FUNCTION_BLOCK DesidratacaoLodo_HMI (* Service Interface Function Block Type *)
  (* Standard: 61499-2 *)
  (* Version 1.2, 21/10/2026, Hidryco, Hidryco, IHM da DesidratacaoLodo 1.2: rodizio e PID nos sub-CATs Revezamento e PID *)
  PACKAGE Hidryco.HidrycoLib;
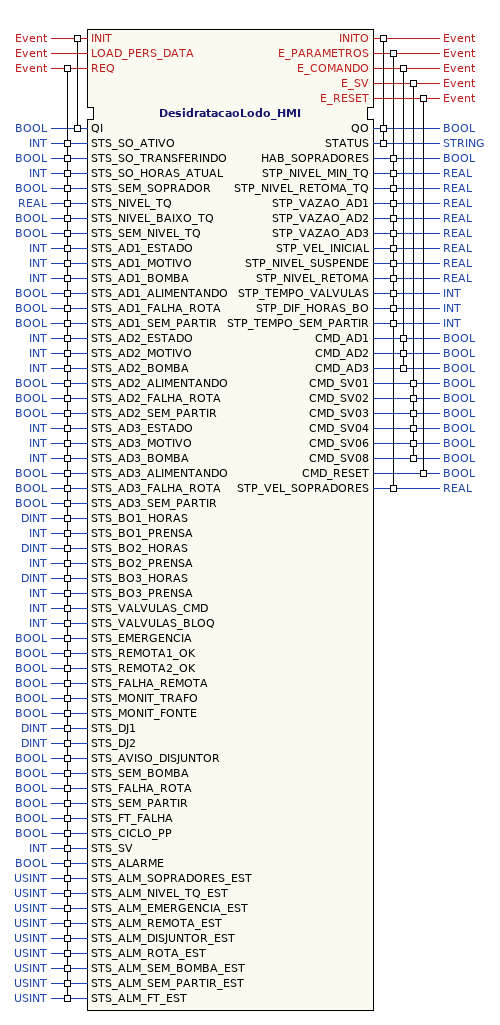
  EVENT_INPUT
    INIT WITH QI;
    LOAD_PERS_DATA; (* Reenvia os parametros persistentes *)
    REQ WITH STS_SO_ATIVO, STS_SO_TRANSFERINDO, STS_SO_HORAS_ATUAL, STS_SEM_SOPRADOR, STS_NIVEL_TQ, STS_NIVEL_BAIXO_TQ, STS_SEM_NIVEL_TQ, STS_AD1_ESTADO, STS_AD1_MOTIVO, STS_AD1_BOMBA, STS_AD1_ALIMENTANDO, STS_AD1_FALHA_ROTA, STS_AD1_SEM_PARTIR, STS_AD2_ESTADO, STS_AD2_MOTIVO, STS_AD2_BOMBA, STS_AD2_ALIMENTANDO, STS_AD2_FALHA_ROTA, STS_AD2_SEM_PARTIR, STS_AD3_ESTADO, STS_AD3_MOTIVO, STS_AD3_BOMBA, STS_AD3_ALIMENTANDO, STS_AD3_FALHA_ROTA, STS_AD3_SEM_PARTIR, STS_BO1_HORAS, STS_BO1_PRENSA, STS_BO2_HORAS, STS_BO2_PRENSA, STS_BO3_HORAS, STS_BO3_PRENSA, STS_VALVULAS_CMD, STS_VALVULAS_BLOQ, STS_EMERGENCIA, STS_REMOTA1_OK, STS_REMOTA2_OK, STS_FALHA_REMOTA, STS_MONIT_TRAFO, STS_MONIT_FONTE, STS_DJ1, STS_DJ2, STS_AVISO_DISJUNTOR, STS_SEM_BOMBA, STS_FALHA_ROTA, STS_SEM_PARTIR, STS_FT_FALHA, STS_CICLO_PP, STS_SV, STS_ALARME, STS_ALM_SOPRADORES_EST, STS_ALM_NIVEL_TQ_EST, STS_ALM_EMERGENCIA_EST, STS_ALM_REMOTA_EST, STS_ALM_DISJUNTOR_EST, STS_ALM_ROTA_EST, STS_ALM_SEM_BOMBA_EST, STS_ALM_SEM_PARTIR_EST, STS_ALM_FT_EST; (* Atualizacao de status *)
  END_EVENT
  EVENT_OUTPUT
    INITO WITH QO, STATUS;
    E_PARAMETROS WITH HAB_SOPRADORES, STP_NIVEL_MIN_TQ, STP_NIVEL_RETOMA_TQ, STP_VAZAO_AD1, STP_VAZAO_AD2, STP_VAZAO_AD3, STP_VEL_INICIAL, STP_NIVEL_SUSPENDE, STP_NIVEL_RETOMA, STP_TEMPO_VALVULAS, STP_DIF_HORAS_BO, STP_TEMPO_SEM_PARTIR, STP_VEL_SOPRADORES;
    E_COMANDO WITH CMD_AD1, CMD_AD2, CMD_AD3;
    E_SV WITH CMD_SV01, CMD_SV02, CMD_SV03, CMD_SV04, CMD_SV06, CMD_SV08;
    E_RESET WITH CMD_RESET;
  END_EVENT
  VAR_INPUT
    QI : BOOL;
    STS_SO_ATIVO : INT; (* Soprador designado: 0 nenhum, 1 SO-01, 2 SO-02 *)
    STS_SO_TRANSFERINDO : BOOL; (* Rodizio em andamento (os dois ligados) *)
    STS_SO_HORAS_ATUAL : INT; (* Horas do soprador atual desde a ultima troca *)
    STS_SEM_SOPRADOR : BOOL; (* Automatico sem nenhum soprador disponivel (risco de sedimentacao) *)
    STS_NIVEL_TQ : REAL; (* Nivel usado no intertravamento (maior entre LIT-01 e LIT-02 validos, %) *)
    STS_NIVEL_BAIXO_TQ : BOOL; (* Tanques de estocagem em nivel baixo: bombas suspensas *)
    STS_SEM_NIVEL_TQ : BOOL; (* LIT-01 e LIT-02 em falha: bombas suspensas *)
    STS_AD1_ESTADO : INT; (* AD-01: 0 parado, 1 abrindo valvulas, 2 partindo bomba, 3 alimentando, 4 suspenso, 5 parando *)
    STS_AD1_MOTIVO : INT; (* AD-01: 0 ok, 1 prensa indisponivel, 2 setpoint zero, 3 sem bomba ou rota, 4 houve falha de rota, 5 emergencia, 6 floculador cheio, 7 tanque baixo, 8 FT em falha, 9 prensa nao partiu *)
    STS_AD1_BOMBA : INT; (* AD-01: bomba em uso (0 nenhuma, 1 a 3 = BO-01 a BO-03) *)
    STS_AD1_ALIMENTANDO : BOOL; (* AD-01 sendo alimentada *)
    STS_AD1_FALHA_ROTA : BOOL; (* AD-01: valvula da rota nao abriu/fechou ou saiu de posicao com a bomba em uso (memorizado; outra rota e tentada) *)
    STS_AD1_SEM_PARTIR : BOOL; (* AD-01 alimentada e a prensa nao partiu no tempo *)
    STS_AD2_ESTADO : INT; (* AD-02: 0 parado, 1 abrindo valvulas, 2 partindo bomba, 3 alimentando, 4 suspenso, 5 parando *)
    STS_AD2_MOTIVO : INT; (* AD-02: 0 ok, 1 prensa indisponivel, 2 setpoint zero, 3 sem bomba ou rota, 4 houve falha de rota, 5 emergencia, 6 floculador cheio, 7 tanque baixo, 8 FT em falha, 9 prensa nao partiu *)
    STS_AD2_BOMBA : INT; (* AD-02: bomba em uso (0 nenhuma, 1 a 3 = BO-01 a BO-03) *)
    STS_AD2_ALIMENTANDO : BOOL; (* AD-02 sendo alimentada *)
    STS_AD2_FALHA_ROTA : BOOL; (* AD-02: valvula da rota nao abriu/fechou ou saiu de posicao com a bomba em uso (memorizado; outra rota e tentada) *)
    STS_AD2_SEM_PARTIR : BOOL; (* AD-02 alimentada e a prensa nao partiu no tempo *)
    STS_AD3_ESTADO : INT; (* AD-03: 0 parado, 1 abrindo valvulas, 2 partindo bomba, 3 alimentando, 4 suspenso, 5 parando *)
    STS_AD3_MOTIVO : INT; (* AD-03: 0 ok, 1 prensa indisponivel, 2 setpoint zero, 3 sem bomba ou rota, 4 houve falha de rota, 5 emergencia, 6 floculador cheio, 7 tanque baixo, 8 FT em falha, 9 prensa nao partiu *)
    STS_AD3_BOMBA : INT; (* AD-03: bomba em uso (0 nenhuma, 1 a 3 = BO-01 a BO-03) *)
    STS_AD3_ALIMENTANDO : BOOL; (* AD-03 sendo alimentada *)
    STS_AD3_FALHA_ROTA : BOOL; (* AD-03: valvula da rota nao abriu/fechou ou saiu de posicao com a bomba em uso (memorizado; outra rota e tentada) *)
    STS_AD3_SEM_PARTIR : BOOL; (* AD-03 alimentada e a prensa nao partiu no tempo *)
    STS_BO1_HORAS : DINT; (* BO-01: horas de operacao (rodizio) *)
    STS_BO1_PRENSA : INT; (* BO-01: prensa atendida (0 nenhuma, 1 a 3) *)
    STS_BO2_HORAS : DINT; (* BO-02: horas de operacao (rodizio) *)
    STS_BO2_PRENSA : INT; (* BO-02: prensa atendida (0 nenhuma, 1 a 3) *)
    STS_BO3_HORAS : DINT; (* BO-03: horas de operacao (rodizio) *)
    STS_BO3_PRENSA : INT; (* BO-03: prensa atendida (0 nenhuma, 1 a 3) *)
    STS_VALVULAS_CMD : INT; (* Valvulas do barrilete comandadas abertas (bit 0 = VA-06 ... bit 7 = VA-13) *)
    STS_VALVULAS_BLOQ : INT; (* Valvulas do barrilete bloqueadas por falha de rota ate o reset (bit 0 = VA-06 ... bit 7 = VA-13) *)
    STS_EMERGENCIA : BOOL; (* Emergencia do PCM LODO acionada *)
    STS_REMOTA1_OK : BOOL; (* Remota 1 do PCE LODO (.135) comunicando *)
    STS_REMOTA2_OK : BOOL; (* Remota 2 do PCE LODO (.136) comunicando *)
    STS_FALHA_REMOTA : BOOL; (* Alguma remota do PCE LODO sem comunicacao *)
    STS_MONIT_TRAFO : BOOL; (* PCM LODO: monitoramento do transformador (%I0.45) *)
    STS_MONIT_FONTE : BOOL; (* PCM LODO: monitoramento da fonte (%I0.51) *)
    STS_DJ1 : DINT; (* Disjuntores ligados, bit 0..15 = PCE, PCM, SO01, SO02, AD01, AD02, AD03, PP01, MN01, MN02, MN03, MN04, MN05, BO01, BO02, BO03 *)
    STS_DJ2 : DINT; (* Disjuntores ligados, bit 0..15 = BR01, BR02, VA01, VA02, VE01, VE02, VA06, VA07, VA08, VA09, VA10, VA11, VA12, VA13, VB03, VB04 *)
    STS_AVISO_DISJUNTOR : BOOL; (* Disjuntor de equipamento existente desligado *)
    STS_SEM_BOMBA : BOOL; (* Prensa pedida sem bomba disponivel *)
    STS_FALHA_ROTA : BOOL; (* Alguma rota de alimentacao com falha de valvula *)
    STS_SEM_PARTIR : BOOL; (* Alguma prensa alimentada sem partir *)
    STS_FT_FALHA : BOOL; (* FT de prensa em falha durante a alimentacao (velocidade mantida) *)
    STS_CICLO_PP : BOOL; (* Ciclo do preparador de polimero ligado pelo automatico *)
    STS_SV : INT; (* Solenoides abertas: bit0 SV-01, bit1 SV-02, bit2 SV-03, bit3 SV-04, bit4 SV-06, bit5 SV-08 *)
    STS_ALARME : BOOL; (* Algum alarme da alimentacao/painel *)
    STS_ALM_SOPRADORES_EST : USINT; (* Estado do ALARM_BIT (0 normal, 1 ativo reconhecido, 2 ativo nao reconhecido, 3 saiu nao reconhecido, 4 ativo e saiu nao reconhecido) *)
    STS_ALM_NIVEL_TQ_EST : USINT; (* Estado do ALARM_BIT (0 normal, 1 ativo reconhecido, 2 ativo nao reconhecido, 3 saiu nao reconhecido, 4 ativo e saiu nao reconhecido) *)
    STS_ALM_EMERGENCIA_EST : USINT; (* Estado do ALARM_BIT (0 normal, 1 ativo reconhecido, 2 ativo nao reconhecido, 3 saiu nao reconhecido, 4 ativo e saiu nao reconhecido) *)
    STS_ALM_REMOTA_EST : USINT; (* Estado do ALARM_BIT (0 normal, 1 ativo reconhecido, 2 ativo nao reconhecido, 3 saiu nao reconhecido, 4 ativo e saiu nao reconhecido) *)
    STS_ALM_DISJUNTOR_EST : USINT; (* Estado do ALARM_BIT (0 normal, 1 ativo reconhecido, 2 ativo nao reconhecido, 3 saiu nao reconhecido, 4 ativo e saiu nao reconhecido) *)
    STS_ALM_ROTA_EST : USINT; (* Estado do ALARM_BIT (0 normal, 1 ativo reconhecido, 2 ativo nao reconhecido, 3 saiu nao reconhecido, 4 ativo e saiu nao reconhecido) *)
    STS_ALM_SEM_BOMBA_EST : USINT; (* Estado do ALARM_BIT (0 normal, 1 ativo reconhecido, 2 ativo nao reconhecido, 3 saiu nao reconhecido, 4 ativo e saiu nao reconhecido) *)
    STS_ALM_SEM_PARTIR_EST : USINT; (* Estado do ALARM_BIT (0 normal, 1 ativo reconhecido, 2 ativo nao reconhecido, 3 saiu nao reconhecido, 4 ativo e saiu nao reconhecido) *)
    STS_ALM_FT_EST : USINT; (* Estado do ALARM_BIT (0 normal, 1 ativo reconhecido, 2 ativo nao reconhecido, 3 saiu nao reconhecido, 4 ativo e saiu nao reconhecido) *)
  END_VAR
  VAR_OUTPUT
    QO : BOOL; (* Event Output Qualifier *)
    STATUS : STRING; (* Service Status *)
    HAB_SOPRADORES : BOOL; (* Sopradores no automatico (um sempre ligado) *)
    STP_NIVEL_MIN_TQ : REAL; (* Nivel minimo dos tanques para as bombas (%); 0 = sem intertravamento *)
    STP_NIVEL_RETOMA_TQ : REAL; (* Nivel dos tanques para retomar as bombas (%) *)
    STP_VAZAO_AD1 : REAL; (* Vazao de lodo da AD-01 (m3/h); 0 = nao alimenta *)
    STP_VAZAO_AD2 : REAL; (* Vazao de lodo da AD-02 (m3/h); 0 = nao alimenta *)
    STP_VAZAO_AD3 : REAL; (* Vazao de lodo da AD-03 (m3/h); 0 = nao alimenta *)
    STP_VEL_INICIAL : REAL; (* Velocidade de partida da bomba (Hz) *)
    STP_NIVEL_SUSPENDE : REAL; (* Floculador: suspende a alimentacao acima deste nivel (%); 0 = desligado *)
    STP_NIVEL_RETOMA : REAL; (* Floculador: retoma abaixo deste nivel (%) *)
    STP_TEMPO_VALVULAS : INT; (* Tempo maximo para abrir as valvulas da rota (s); 0 = sem limite *)
    STP_DIF_HORAS_BO : INT; (* Rodizio das bombas: BO-02 assume quando a titular tem estas horas a mais; 0 = sem rodizio *)
    STP_TEMPO_SEM_PARTIR : INT; (* Aviso se a prensa nao partir com alimentacao (min); 0 = desligado *)
    CMD_AD1 : BOOL; (* Desaguamento ligado na AD-01 (nao persistente: apos reinicio do CLP o operador religa) *)
    CMD_AD2 : BOOL; (* Desaguamento ligado na AD-02 (nao persistente: apos reinicio do CLP o operador religa) *)
    CMD_AD3 : BOOL; (* Desaguamento ligado na AD-03 (nao persistente: apos reinicio do CLP o operador religa) *)
    CMD_SV01 : BOOL; (* Abre a 900-SV-01 (manual) *)
    CMD_SV02 : BOOL; (* Abre a 900-SV-02 (manual) *)
    CMD_SV03 : BOOL; (* Abre a 900-SV-03 (manual) *)
    CMD_SV04 : BOOL; (* Abre a 900-SV-04 (manual) *)
    CMD_SV06 : BOOL; (* Abre a 900-SV-06 (manual) *)
    CMD_SV08 : BOOL; (* Abre a 900-SV-08 (manual) *)
    CMD_RESET : BOOL; (* Reconhece os alarmes da fase solida *)
    STP_VEL_SOPRADORES : REAL; (* Velocidade dos sopradores no automatico (Hz) *)
  END_VAR
  SERVICE /
    SEQUENCE 
    END_SEQUENCE
  END_SERVICE
END_FUNCTION_BLOCK
